PROGRAM MAIN
VAR
    Clock         : TaskClock(CycleTime := LTIME#10MS);

    // Filling station: every candidate is declared; the routers choose
    RealTankValve  : SolenoidValve(Output := GVL_Io.TankValveCoil,
                                   OpenFeedback := GVL_Io.TankValveOpen,
                                   FaultDelay := T#2S);
    SimTankValve   : SimulatedValve(Name := 'Tank valve', Clock := Clock, TravelTime := LTIME#400MS);
    TankValve      : FillValveRouter(Name := 'Tank valve', Source := GVL_Site.TankValveSource,
                                     FinalHardware := RealTankValve, SimilarHardware := 0,
                                     Simulation := SimTankValve, Test := 0);

    RealDrainValve : SolenoidValve(Output := GVL_Io.DrainValveCoil,
                                   OpenFeedback := GVL_Io.DrainValveOpen,
                                   FaultDelay := T#2S);
    SimDrainValve  : SimulatedValve(Name := 'Drain valve', Clock := Clock, TravelTime := LTIME#400MS);
    DrainValve     : FillValveRouter(Name := 'Drain valve', Source := GVL_Site.DrainValveSource,
                                     FinalHardware := RealDrainValve, SimilarHardware := 0,
                                     Simulation := SimDrainValve, Test := 0);

    SimTank        : TankModel(Inflow := TankValve, Outflow := DrainValve, Clock := Clock,
                               FillRate := 20.0, DrainRate := 25.0, StartLevel := 0.0);
    RealLevel      : FieldbusLevelSensor(FieldbusLevel := GVL_Io.TankLevel,
                                         IsCommunicationOk := GVL_Io.TankSensorOk,
                                         TankHeight := 300.0);          // the dosing tank, mm
    TankLevel      : LevelSensorRouter(Name := 'Tank level', Source := GVL_Site.TankLevelSource,
                                       FinalHardware := RealLevel, SimilarHardware := 0,
                                       Simulation := SimTank, Test := 0);

    // Pick-and-place station
    RealLift       : SingleSolenoidCylinder(Name := 'Lift', MoveTimeout := T#1S,
                                            Solenoid := GVL_Io.LiftValve,
                                            ExtendedSensor := GVL_Io.LiftDown,
                                            RetractedSensor := GVL_Io.LiftUp);
    SimLift        : SimulatedActuator(Name := 'Lift', MoveTimeout := T#1S, TravelTime := T#400MS);
    LiftCylinder   : ActuatorRouter(Name := 'Lift', Source := GVL_Site.LiftSource,
                                    FinalHardware := RealLift, SimilarHardware := 0,
                                    Simulation := SimLift, Test := 0);

    RealSlide      : DoubleSolenoidCylinder(Name := 'Slide', MoveTimeout := T#2S,
                                            ExtendCoil := GVL_Io.SlideOutCoil,
                                            RetractCoil := GVL_Io.SlideInCoil,
                                            ExtendedSensor := GVL_Io.SlideOut,
                                            RetractedSensor := GVL_Io.SlideIn);
    SimSlide       : SimulatedActuator(Name := 'Slide', MoveTimeout := T#2S, TravelTime := T#800MS);
    SlideCylinder  : ActuatorRouter(Name := 'Slide', Source := GVL_Site.SlideSource,
                                    FinalHardware := RealSlide, SimilarHardware := 0,
                                    Simulation := SimSlide, Test := 0);

    RealGripper    : Gripper(Name := 'Gripper', MoveTimeout := T#500MS,
                             Solenoid := GVL_Io.GripperValve,
                             ExtendedSensor := GVL_Io.GripperClosed,
                             RetractedSensor := GVL_Io.GripperOpen);
    SimGripper     : SimulatedActuator(Name := 'Gripper', MoveTimeout := T#500MS, TravelTime := T#150MS);
    PartGripper    : ActuatorRouter(Name := 'Gripper', Source := GVL_Site.GripperSource,
                                    FinalHardware := RealGripper, SimilarHardware := 0,
                                    Simulation := SimGripper, Test := 0);

    // The operations, unchanged from their pages
    TankFill       : FillSequence(LevelSensor := TankLevel, FillValve := TankValve);
    Dose           : DrainTankCommand(DrainValve := DrainValve, Level := TankLevel,
                                      Clock := Clock, Timeout := LTIME#30S);
    PickPlace      : PickAndPlaceSequence(Lift := LiftCylinder, Slide := SlideCylinder,
                                          Gripper := PartGripper);

    // The tree
    Sources        : SimulationCheck(IsOnMachine := GVL_Site.IsOnMachine);
    Filling        : FillingModule(Name := 'Filling', Fill := TankFill, Dose := Dose);
    PickAndPlace   : PickAndPlaceModule(Name := 'Pick and place', Sequence := PickPlace);
    Line           : LineModule(Name := 'Line 1', Filler := Filling, Transfer := PickAndPlace);

    StartEdge      : R_TRIG;
    StopEdge       : R_TRIG;
    ResetEdge      : R_TRIG;
    Wired          : BOOL;
    WiredOk        : BOOL;
END_VAR

// Build the tree once, and tell the check where every device comes from
IF NOT Wired THEN
    Wired := TRUE;
    WiredOk := Filling.AddChild(Child := TankValve);
    WiredOk := Filling.AddChild(Child := DrainValve) AND WiredOk;
    WiredOk := PickAndPlace.AddChild(Child := LiftCylinder) AND WiredOk;
    WiredOk := PickAndPlace.AddChild(Child := SlideCylinder) AND WiredOk;
    WiredOk := PickAndPlace.AddChild(Child := PartGripper) AND WiredOk;
    WiredOk := Line.AddChild(Child := Sources) AND WiredOk;
    WiredOk := Line.AddChild(Child := Filling) AND WiredOk;
    WiredOk := Line.AddChild(Child := PickAndPlace) AND WiredOk;

    WiredOk := Sources.AddDevice(Name := TankValve.Name, Source := TankValve.Source) AND WiredOk;
    WiredOk := Sources.AddDevice(Name := DrainValve.Name, Source := DrainValve.Source) AND WiredOk;
    WiredOk := Sources.AddDevice(Name := TankLevel.Name, Source := TankLevel.Source) AND WiredOk;
    WiredOk := Sources.AddDevice(Name := LiftCylinder.Name, Source := LiftCylinder.Source) AND WiredOk;
    WiredOk := Sources.AddDevice(Name := SlideCylinder.Name, Source := SlideCylinder.Source) AND WiredOk;
    WiredOk := Sources.AddDevice(Name := PartGripper.Name, Source := PartGripper.Source) AND WiredOk;
    GVL_Hmi.NotFinalDevices := Sources.NotFinalDevices;
END_IF

// Failure hooks act only on a simulated device
IF TankValve.Source = E_DeviceSource.Simulation THEN
    SimTankValve.SetStuck(IsStuck := GVL_Sim.TankValveStuck);
END_IF
IF DrainValve.Source = E_DeviceSource.Simulation THEN
    SimDrainValve.SetStuck(IsStuck := GVL_Sim.DrainValveStuck);
END_IF
IF LiftCylinder.Source = E_DeviceSource.Simulation THEN
    SimLift.SetStuck(IsStuck := GVL_Sim.LiftStuck);
END_IF
IF SlideCylinder.Source = E_DeviceSource.Simulation THEN
    SimSlide.SetStuck(IsStuck := GVL_Sim.SlideStuck);
END_IF
IF PartGripper.Source = E_DeviceSource.Simulation THEN
    SimGripper.SetStuck(IsStuck := GVL_Sim.GripperStuck);
END_IF

// Operator commands
StartEdge(CLK := GVL_Hmi.StartButton);
StopEdge(CLK := GVL_Hmi.StopButton);
ResetEdge(CLK := GVL_Hmi.ResetButton);
IF StartEdge.Q AND WiredOk THEN
    Line.Start();
END_IF
IF StopEdge.Q THEN
    Line.Stop();
END_IF
IF ResetEdge.Q THEN
    Line.Reset();
END_IF

Clock.CyclicLogic();                            // first: everything below reads its time
TankLevel.CyclicLogic();                        // runs the tank model only when it's the chosen level
Line.CyclicLogic();                             // the line, then each station, then its devices

GVL_Hmi.LineState := Line.State;
GVL_Hmi.IsStopping := Line.IsStopping;
GVL_Hmi.FaultText := Line.FaultText;

END_PROGRAM

(* stored: Version 1.1.0.1, ProductVersion 3.1.4026.0
   POU MAIN: Id {7c92886d-c7ab-4116-ba27-be0f4b76e777}, SpecialFunc None *)
